FUNCTION_BLOCK INIT_OFF (* E_TRIG Counterpart, erweitert um ein eigenstaendiges INIT_OFF/INITO_OFF Pass-Through (EInitOff) *)
  (* Standard: 61131-3; Classification: standard boolean function; Description: Copyright (c) 2026 Meisterschulen am Ostbahnhof This program and the accompanying materials are made available under the terms of the Eclipse Public License 2.0 which is available at https://www.eclipse.org/legal/epl-2.0/ SPDX-License-Identifier: EPL-2.0 *)
  (* Version 1.0, 2026-10-11, Franz Höpfinger, Meisterschulen am Ostbahnhof, initial API and implementation and/or initial documentation. Basiert auf dem INIT.fbt Pass-Through-Muster, ergaenzt um einen zweiten, unabhaengigen Init-Kanal INIT_OFF/INITO_OFF (EInitOff). Pendant zu INIT_ON.fbt. *)
  PACKAGE events::init;
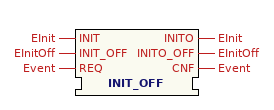
  EVENT_INPUT
    INIT : EInit; (* Initialization Request *)
    INIT_OFF : EInitOff; (* Initialization Request, eigener Kanal unabhaengig von INIT *)
    REQ; (* Service Request *)
  END_EVENT
  EVENT_OUTPUT
    INITO : EInit; (* Initialization Confirm *)
    INITO_OFF : EInitOff; (* Initialization Confirm, eigener Kanal unabhaengig von INITO *)
    CNF; (* Confirmation of Requested Service *)
  END_EVENT
  EVENT_CONNECTIONS
    INIT TO INITO;
    REQ TO CNF;
    INIT_OFF TO INITO_OFF;
  END_CONNECTIONS
END_FUNCTION_BLOCK
